{attribute 'no_assign'}
FUNCTION_BLOCK FB_DO_WTURBINE_LD0_WPPD1_DevSt EXTENDS FB_AcsiCommonDataClass
VAR_INPUT
	st_: FB_DO_WTURBINE_LD0_WPPD1_DevSt_st := (sObjectName:='st', sClass:='ENS', bLinkResult:=THIS^.AddDataToContainer(ipData:=st_));
END_VAR
VAR
END_VAR

END_FUNCTION_BLOCK

(* stored: Version 1.1.0.1
   POU FB_DO_WTURBINE_LD0_WPPD1_DevSt: Id {048aabed-4892-4300-8203-b2d8ef23180a}, SpecialFunc None *)
